{region 'Documentation'}
(*!
<summary>Withholds CompleteAbort and verifies timeout finalization with the latched Abort timeout flag.</summary>
*)
{endregion}
FUNCTION_BLOCK Test_LifecycleAbortTimeout EXTENDS TestCaseLifecycleTestBase

SUPER^();

{region 'Documentation'}
(*!
<summary>Defines explicit exceptional-path stimuli and contract-derived observations.</summary>
*)
{endregion}
METHOD PROTECTED ConfigureScenario
// Exercise the real cyclic timer; these checkpoints check the timeout path and retained flag,
// not an exact elapsed-time boundary. The outer Test Case timeout bounds a missing transition.
FSubjectPreparationCount := 0;
FSubjectTestCount := 1;
FStepCount := 12;
FSubjectConfig.AbortTimeout := T#50ms;

{region "01 - Reset to Idle"}
// Establish Idle through the parent Reset request; both child results must be cleared.
FSteps[1].RequestReset := TRUE;
FSteps[1].ExpectedState := E_State.Idle;
FSteps[1].ExpectedResult := E_Result.NotEvaluated;
FSteps[1].ExpectedReady := TRUE;
FSteps[1].ExpectedPassedCount := 0;
FSteps[1].ExpectedFailedCount := 0;
FSteps[1].ExpectedHookCount := 6;
FSteps[1].ExpectedHooks[1].Hook := E_LifecycleHook.Reset;
FSteps[1].ExpectedHooks[1].State := E_State.Reset;
FSteps[1].ExpectedHooks[1].Enabled := TRUE;
FSteps[1].ExpectedHooks[2].Hook := E_LifecycleHook.Abort;
FSteps[1].ExpectedHooks[2].State := E_State.Idle;
FSteps[1].ExpectedHooks[2].Enabled := FALSE;
FSteps[1].ExpectedHooks[3].Hook := E_LifecycleHook.Preparations;
FSteps[1].ExpectedHooks[3].State := E_State.Idle;
FSteps[1].ExpectedHooks[3].Enabled := FALSE;
FSteps[1].ExpectedHooks[4].Hook := E_LifecycleHook.Tests;
FSteps[1].ExpectedHooks[4].State := E_State.Idle;
FSteps[1].ExpectedHooks[4].Enabled := FALSE;
FSteps[1].ExpectedHooks[5].Hook := E_LifecycleHook.Assertions;
FSteps[1].ExpectedHooks[5].State := E_State.Idle;
FSteps[1].ExpectedHooks[5].Enabled := FALSE;
FSteps[1].ExpectedHooks[6].Hook := E_LifecycleHook.Aggregate;
FSteps[1].ExpectedHooks[6].State := E_State.Idle;
FSteps[1].ExpectedHooks[6].Enabled := TRUE;
{endregion}

{region "02 - Accept Start"}
// Accept Start into Starting; processing and Assertion evaluation are not active yet.
FSteps[2].RequestStart := TRUE;
FSteps[2].ExpectedState := E_State.Starting;
FSteps[2].ExpectedResult := E_Result.NotEvaluated;
FSteps[2].ExpectedReady := FALSE;
FSteps[2].ExpectedPassedCount := 0;
FSteps[2].ExpectedFailedCount := 0;
FSteps[2].ExpectedHookCount := 5;
FSteps[2].ExpectedHooks[1].Hook := E_LifecycleHook.Abort;
FSteps[2].ExpectedHooks[1].State := E_State.Starting;
FSteps[2].ExpectedHooks[1].Enabled := FALSE;
FSteps[2].ExpectedHooks[2].Hook := E_LifecycleHook.Preparations;
FSteps[2].ExpectedHooks[2].State := E_State.Starting;
FSteps[2].ExpectedHooks[2].Enabled := FALSE;
FSteps[2].ExpectedHooks[3].Hook := E_LifecycleHook.Tests;
FSteps[2].ExpectedHooks[3].State := E_State.Starting;
FSteps[2].ExpectedHooks[3].Enabled := FALSE;
FSteps[2].ExpectedHooks[4].Hook := E_LifecycleHook.Assertions;
FSteps[2].ExpectedHooks[4].State := E_State.Starting;
FSteps[2].ExpectedHooks[4].Enabled := FALSE;
FSteps[2].ExpectedHooks[5].Hook := E_LifecycleHook.Aggregate;
FSteps[2].ExpectedHooks[5].State := E_State.Starting;
FSteps[2].ExpectedHooks[5].Enabled := TRUE;
{endregion}

{region "03 - Enter Running"}
// Enter Running and evaluate both children; owner Result stays NotEvaluated until finalization.
FSteps[3].ExpectedState := E_State.Running;
FSteps[3].ExpectedResult := E_Result.NotEvaluated;
FSteps[3].ExpectedReady := FALSE;
FSteps[3].ExpectedPassedCount := 2;
FSteps[3].ExpectedFailedCount := 0;
FSteps[3].ExpectedHookCount := 5;
FSteps[3].ExpectedHooks[1].Hook := E_LifecycleHook.Abort;
FSteps[3].ExpectedHooks[1].State := E_State.Running;
FSteps[3].ExpectedHooks[1].Enabled := FALSE;
FSteps[3].ExpectedHooks[2].Hook := E_LifecycleHook.Preparations;
FSteps[3].ExpectedHooks[2].State := E_State.Running;
FSteps[3].ExpectedHooks[2].Enabled := FALSE;
FSteps[3].ExpectedHooks[3].Hook := E_LifecycleHook.Tests;
FSteps[3].ExpectedHooks[3].State := E_State.Running;
FSteps[3].ExpectedHooks[3].Enabled := TRUE;
FSteps[3].ExpectedHooks[4].Hook := E_LifecycleHook.Assertions;
FSteps[3].ExpectedHooks[4].State := E_State.Running;
FSteps[3].ExpectedHooks[4].Enabled := TRUE;
FSteps[3].ExpectedHooks[5].Hook := E_LifecycleHook.Aggregate;
FSteps[3].ExpectedHooks[5].State := E_State.Running;
FSteps[3].ExpectedHooks[5].Enabled := TRUE;
{endregion}

{region "04 - Request Abort and hold acknowledgement"}
// Request Abort once and withhold cleanup acknowledgement.
FSteps[4].RequestAbort := TRUE;
FSteps[4].AbortCompleted := FALSE;
FSteps[4].ExpectedState := E_State.Aborting;
FSteps[4].ExpectedResult := E_Result.Abort;
FSteps[4].ExpectedReady := FALSE;
FSteps[4].ExpectedPassedCount := 2;
FSteps[4].ExpectedFailedCount := 0;
FSteps[4].ExpectedHookCount := 5;
FSteps[4].ExpectedHooks[1].Hook := E_LifecycleHook.Abort;
FSteps[4].ExpectedHooks[1].State := E_State.Aborting;
FSteps[4].ExpectedHooks[1].Enabled := TRUE;
FSteps[4].ExpectedHooks[2].Hook := E_LifecycleHook.Preparations;
FSteps[4].ExpectedHooks[2].State := E_State.Aborting;
FSteps[4].ExpectedHooks[2].Enabled := FALSE;
FSteps[4].ExpectedHooks[3].Hook := E_LifecycleHook.Tests;
FSteps[4].ExpectedHooks[3].State := E_State.Aborting;
FSteps[4].ExpectedHooks[3].Enabled := FALSE;
FSteps[4].ExpectedHooks[4].Hook := E_LifecycleHook.Assertions;
FSteps[4].ExpectedHooks[4].State := E_State.Aborting;
FSteps[4].ExpectedHooks[4].Enabled := FALSE;
FSteps[4].ExpectedHooks[5].Hook := E_LifecycleHook.Aggregate;
FSteps[4].ExpectedHooks[5].State := E_State.Aborting;
FSteps[4].ExpectedHooks[5].Enabled := TRUE;
{endregion}

{region "05 - Wait for Abort timeout"}
// Keep cleanup open while repeating this checkpoint in Aborting.
// Timeout forces Completing with Error even though the implementation never acknowledges Abort.
FSteps[5].WaitForTransition := TRUE;
FSteps[5].WaitingState := E_State.Aborting;
FSteps[5].AbortCompleted := FALSE;
FSteps[5].ExpectedAbortTimeout := TRUE;
FSteps[5].ExpectedState := E_State.Completing;
FSteps[5].ExpectedResult := E_Result.Error;
FSteps[5].ExpectedReady := FALSE;
FSteps[5].ExpectedPassedCount := 2;
FSteps[5].ExpectedFailedCount := 0;
FSteps[5].ExpectedHookCount := 5;
FSteps[5].ExpectedHooks[1].Hook := E_LifecycleHook.Abort;
FSteps[5].ExpectedHooks[1].State := E_State.Completing;
FSteps[5].ExpectedHooks[1].Enabled := FALSE;
FSteps[5].ExpectedHooks[2].Hook := E_LifecycleHook.Preparations;
FSteps[5].ExpectedHooks[2].State := E_State.Completing;
FSteps[5].ExpectedHooks[2].Enabled := FALSE;
FSteps[5].ExpectedHooks[3].Hook := E_LifecycleHook.Tests;
FSteps[5].ExpectedHooks[3].State := E_State.Completing;
FSteps[5].ExpectedHooks[3].Enabled := FALSE;
FSteps[5].ExpectedHooks[4].Hook := E_LifecycleHook.Assertions;
FSteps[5].ExpectedHooks[4].State := E_State.Completing;
FSteps[5].ExpectedHooks[4].Enabled := FALSE;
FSteps[5].ExpectedHooks[5].Hook := E_LifecycleHook.Aggregate;
FSteps[5].ExpectedHooks[5].State := E_State.Completing;
FSteps[5].ExpectedHooks[5].Enabled := TRUE;
{endregion}

{region "06 - Retain timeout at completion"}
// Reach Completed and retain the Abort-timeout diagnostic.
FSteps[6].ExpectedAbortTimeout := TRUE;
FSteps[6].ExpectedState := E_State.Completed;
FSteps[6].ExpectedResult := E_Result.Error;
FSteps[6].ExpectedReady := FALSE;
FSteps[6].ExpectedPassedCount := 2;
FSteps[6].ExpectedFailedCount := 0;
FSteps[6].ExpectedHookCount := 1;
FSteps[6].ExpectedHooks[1].Hook := E_LifecycleHook.Aggregate;
FSteps[6].ExpectedHooks[1].State := E_State.Completed;
FSteps[6].ExpectedHooks[1].Enabled := TRUE;
{endregion}

{region "07 - Reset clears held timeout and result"}
FSteps[7].ExpectedState := E_State.Idle;
FSteps[7].ExpectedResult := E_Result.NotEvaluated;
FSteps[7].ExpectedReady := TRUE;
FSteps[7].ExpectedPassedCount := 0;
FSteps[7].ExpectedFailedCount := 0;
FSteps[7].CheckFinalization := TRUE;
FSteps[7].ExpectedFinalizationCount := 1;
FSteps[7].ExpectedCompletionCount := 1;
FSteps[7].ExpectedFinalResult := E_Result.Error;
FSteps[7].RequestReset := TRUE;
FSteps[7].PreparationTargetReached := TRUE;
FSteps[7].ExpectRuntimeCleared := TRUE;
FSteps[7].ExpectedHookCount := 6;
FSteps[7].ExpectedHooks[1].Hook := E_LifecycleHook.Reset;
FSteps[7].ExpectedHooks[1].State := E_State.Reset;
FSteps[7].ExpectedHooks[1].Enabled := TRUE;
FSteps[7].ExpectedHooks[2].Hook := E_LifecycleHook.Abort;
FSteps[7].ExpectedHooks[2].State := E_State.Idle;
FSteps[7].ExpectedHooks[2].Enabled := FALSE;
FSteps[7].ExpectedHooks[3].Hook := E_LifecycleHook.Preparations;
FSteps[7].ExpectedHooks[3].State := E_State.Idle;
FSteps[7].ExpectedHooks[3].Enabled := FALSE;
FSteps[7].ExpectedHooks[4].Hook := E_LifecycleHook.Tests;
FSteps[7].ExpectedHooks[4].State := E_State.Idle;
FSteps[7].ExpectedHooks[4].Enabled := FALSE;
FSteps[7].ExpectedHooks[5].Hook := E_LifecycleHook.Assertions;
FSteps[7].ExpectedHooks[5].State := E_State.Idle;
FSteps[7].ExpectedHooks[5].Enabled := FALSE;
FSteps[7].ExpectedHooks[6].Hook := E_LifecycleHook.Aggregate;
FSteps[7].ExpectedHooks[6].State := E_State.Idle;
FSteps[7].ExpectedHooks[6].Enabled := TRUE;
{endregion}

{region "08 - Start after timeout recovery"}
FSteps[8].ExpectedState := E_State.Starting;
FSteps[8].ExpectedResult := E_Result.NotEvaluated;
FSteps[8].ExpectedReady := FALSE;
FSteps[8].ExpectedPassedCount := 0;
FSteps[8].ExpectedFailedCount := 0;
FSteps[8].CheckFinalization := TRUE;
FSteps[8].ExpectedFinalizationCount := 1;
FSteps[8].ExpectedCompletionCount := 1;
FSteps[8].ExpectedFinalResult := E_Result.Error;
FSteps[8].RequestStart := TRUE;
FSteps[8].PreparationTargetReached := TRUE;
FSteps[8].ExpectedHookCount := 5;
FSteps[8].ExpectedHooks[1].Hook := E_LifecycleHook.Abort;
FSteps[8].ExpectedHooks[1].State := E_State.Starting;
FSteps[8].ExpectedHooks[1].Enabled := FALSE;
FSteps[8].ExpectedHooks[2].Hook := E_LifecycleHook.Preparations;
FSteps[8].ExpectedHooks[2].State := E_State.Starting;
FSteps[8].ExpectedHooks[2].Enabled := FALSE;
FSteps[8].ExpectedHooks[3].Hook := E_LifecycleHook.Tests;
FSteps[8].ExpectedHooks[3].State := E_State.Starting;
FSteps[8].ExpectedHooks[3].Enabled := FALSE;
FSteps[8].ExpectedHooks[4].Hook := E_LifecycleHook.Assertions;
FSteps[8].ExpectedHooks[4].State := E_State.Starting;
FSteps[8].ExpectedHooks[4].Enabled := FALSE;
FSteps[8].ExpectedHooks[5].Hook := E_LifecycleHook.Aggregate;
FSteps[8].ExpectedHooks[5].State := E_State.Starting;
FSteps[8].ExpectedHooks[5].Enabled := TRUE;
{endregion}

{region "09 - Execute without previous timeout flags"}
FSteps[9].ExpectedState := E_State.Running;
FSteps[9].ExpectedResult := E_Result.NotEvaluated;
FSteps[9].ExpectedReady := FALSE;
FSteps[9].ExpectedPassedCount := 2;
FSteps[9].ExpectedFailedCount := 0;
FSteps[9].CheckFinalization := TRUE;
FSteps[9].ExpectedFinalizationCount := 1;
FSteps[9].ExpectedCompletionCount := 1;
FSteps[9].ExpectedFinalResult := E_Result.Error;
FSteps[9].ExpectedHookCount := 5;
FSteps[9].ExpectedHooks[1].Hook := E_LifecycleHook.Abort;
FSteps[9].ExpectedHooks[1].State := E_State.Running;
FSteps[9].ExpectedHooks[1].Enabled := FALSE;
FSteps[9].ExpectedHooks[2].Hook := E_LifecycleHook.Preparations;
FSteps[9].ExpectedHooks[2].State := E_State.Running;
FSteps[9].ExpectedHooks[2].Enabled := FALSE;
FSteps[9].ExpectedHooks[3].Hook := E_LifecycleHook.Tests;
FSteps[9].ExpectedHooks[3].State := E_State.Running;
FSteps[9].ExpectedHooks[3].Enabled := TRUE;
FSteps[9].ExpectedHooks[4].Hook := E_LifecycleHook.Assertions;
FSteps[9].ExpectedHooks[4].State := E_State.Running;
FSteps[9].ExpectedHooks[4].Enabled := TRUE;
FSteps[9].ExpectedHooks[5].Hook := E_LifecycleHook.Aggregate;
FSteps[9].ExpectedHooks[5].State := E_State.Running;
FSteps[9].ExpectedHooks[5].Enabled := TRUE;
{endregion}

{region "10 - Finalize the recovered run"}
FSteps[10].ExpectedState := E_State.Completing;
FSteps[10].ExpectedResult := E_Result.Passed;
FSteps[10].ExpectedReady := FALSE;
FSteps[10].ExpectedPassedCount := 2;
FSteps[10].ExpectedFailedCount := 0;
FSteps[10].FinishTests := TRUE;
FSteps[10].CheckFinalization := TRUE;
FSteps[10].ExpectedFinalizationCount := 2;
FSteps[10].ExpectedCompletionCount := 1;
FSteps[10].ExpectedFinalResult := E_Result.Passed;
FSteps[10].ExpectedHookCount := 5;
FSteps[10].ExpectedHooks[1].Hook := E_LifecycleHook.Abort;
FSteps[10].ExpectedHooks[1].State := E_State.Running;
FSteps[10].ExpectedHooks[1].Enabled := FALSE;
FSteps[10].ExpectedHooks[2].Hook := E_LifecycleHook.Preparations;
FSteps[10].ExpectedHooks[2].State := E_State.Running;
FSteps[10].ExpectedHooks[2].Enabled := FALSE;
FSteps[10].ExpectedHooks[3].Hook := E_LifecycleHook.Tests;
FSteps[10].ExpectedHooks[3].State := E_State.Running;
FSteps[10].ExpectedHooks[3].Enabled := TRUE;
FSteps[10].ExpectedHooks[4].Hook := E_LifecycleHook.Assertions;
FSteps[10].ExpectedHooks[4].State := E_State.Completing;
FSteps[10].ExpectedHooks[4].Enabled := FALSE;
FSteps[10].ExpectedHooks[5].Hook := E_LifecycleHook.Aggregate;
FSteps[10].ExpectedHooks[5].State := E_State.Completing;
FSteps[10].ExpectedHooks[5].Enabled := TRUE;
{endregion}

{region "11 - Complete the recovered run"}
FSteps[11].ExpectedState := E_State.Completed;
FSteps[11].ExpectedResult := E_Result.Passed;
FSteps[11].ExpectedReady := FALSE;
FSteps[11].ExpectedPassedCount := 2;
FSteps[11].ExpectedFailedCount := 0;
FSteps[11].ExpectRuntimeHeld := TRUE;
FSteps[11].CheckFinalization := TRUE;
FSteps[11].ExpectedFinalizationCount := 2;
FSteps[11].ExpectedCompletionCount := 2;
FSteps[11].ExpectedFinalResult := E_Result.Passed;
FSteps[11].ExpectedHookCount := 1;
FSteps[11].ExpectedHooks[1].Hook := E_LifecycleHook.Aggregate;
FSteps[11].ExpectedHooks[1].State := E_State.Completed;
FSteps[11].ExpectedHooks[1].Enabled := TRUE;
{endregion}

{region "12 - Hold the recovered completion without new events"}
FSteps[12].ExpectedState := E_State.Completed;
FSteps[12].ExpectedResult := E_Result.Passed;
FSteps[12].ExpectedReady := FALSE;
FSteps[12].ExpectedPassedCount := 2;
FSteps[12].ExpectedFailedCount := 0;
FSteps[12].ExpectQuietCall := TRUE;
FSteps[12].ExpectRuntimeHeld := TRUE;
FSteps[12].CheckFinalization := TRUE;
FSteps[12].ExpectedFinalizationCount := 2;
FSteps[12].ExpectedCompletionCount := 2;
FSteps[12].ExpectedFinalResult := E_Result.Passed;
FSteps[12].ExpectedHookCount := 1;
FSteps[12].ExpectedHooks[1].Hook := E_LifecycleHook.Aggregate;
FSteps[12].ExpectedHooks[1].State := E_State.Completed;
FSteps[12].ExpectedHooks[1].Enabled := TRUE;
{endregion}
END_METHOD

END_FUNCTION_BLOCK

(* stored: Version 1.1.0.1
   POU Test_LifecycleAbortTimeout: Id {fd3790d8-7519-4c3a-9fe3-7cb135f093ca}, SpecialFunc None
   Folder Internal: Id {205df96b-198f-4c0a-9666-4cb363311495}
   Method ConfigureScenario: Id {71605b52-2ae4-4dda-b764-08935667fe19} *)
